FUNCTION "ROLL_PB25" : Void
{ S7_Optimized_Access := 'TRUE' }
VERSION : 0.1
VAR_TEMP
    r : Bool;
    a1 : Word;
    a2 : Word;
    activeDataBlock : Int;
    comparisonResults : Array[0..14] of Bool;
END_VAR
BEGIN
    #r := FALSE;
    #a1 := W#16#0000;
    #a2 := W#16#0000;
    #activeDataBlock := 0;
    // PB25, STEP 5 network 1
    #activeDataBlock := 15;
    // PB25, STEP 5 network 2
    #a2 := #a1;
    #a1 := "ROLL_GetM"(FirstByte := 5, Width := 8);
    #a2 := #a1;
    #a1 := W#16#0000;
    #comparisonResults[0] := (WORD_TO_INT(#a2) <> WORD_TO_INT(#a1));
    #r := #comparisonResults[0];
    "ROLL_State".M[87, 0] := #r;
    // PB25, STEP 5 network 3
    #a2 := #a1;
    #a1 := "ROLL_GetM"(FirstByte := 6, Width := 8);
    #a2 := #a1;
    #a1 := W#16#0000;
    #comparisonResults[1] := (WORD_TO_INT(#a2) <> WORD_TO_INT(#a1));
    #r := #comparisonResults[1];
    "ROLL_State".M[87, 1] := #r;
    // PB25, STEP 5 network 4
    #a2 := #a1;
    #a1 := "ROLL_GetM"(FirstByte := 7, Width := 8);
    #a2 := #a1;
    #a1 := W#16#0000;
    #comparisonResults[2] := (WORD_TO_INT(#a2) <> WORD_TO_INT(#a1));
    #r := #comparisonResults[2];
    "ROLL_State".M[87, 2] := #r;
    // PB25, STEP 5 network 5
    #a2 := #a1;
    #a1 := "ROLL_GetM"(FirstByte := 8, Width := 8);
    #a2 := #a1;
    #a1 := W#16#0000;
    #comparisonResults[3] := (WORD_TO_INT(#a2) <> WORD_TO_INT(#a1));
    #r := #comparisonResults[3];
    "ROLL_State".M[87, 3] := #r;
    // PB25, STEP 5 network 6
    #a2 := #a1;
    #a1 := "ROLL_GetM"(FirstByte := 9, Width := 8);
    #a2 := #a1;
    #a1 := W#16#0000;
    #comparisonResults[4] := (WORD_TO_INT(#a2) <> WORD_TO_INT(#a1));
    #r := #comparisonResults[4];
    "ROLL_State".M[87, 4] := #r;
    // PB25, STEP 5 network 7
    #a2 := #a1;
    #a1 := "ROLL_GetM"(FirstByte := 10, Width := 8);
    #a2 := #a1;
    #a1 := W#16#0000;
    #comparisonResults[5] := (WORD_TO_INT(#a2) <> WORD_TO_INT(#a1));
    #r := #comparisonResults[5];
    "ROLL_State".M[87, 5] := #r;
    // PB25, STEP 5 network 8
    #a2 := #a1;
    #a1 := "ROLL_GetM"(FirstByte := 11, Width := 8);
    #a2 := #a1;
    #a1 := W#16#0000;
    #comparisonResults[6] := (WORD_TO_INT(#a2) <> WORD_TO_INT(#a1));
    #r := #comparisonResults[6];
    "ROLL_State".M[87, 6] := #r;
    // PB25, STEP 5 network 9
    #a2 := #a1;
    #a1 := "ROLL_GetM"(FirstByte := 12, Width := 8);
    #a2 := #a1;
    #a1 := W#16#0000;
    #comparisonResults[7] := (WORD_TO_INT(#a2) <> WORD_TO_INT(#a1));
    #r := #comparisonResults[7];
    "ROLL_State".M[87, 7] := #r;
    // PB25, STEP 5 network 10
    #a2 := #a1;
    #a1 := "ROLL_GetM"(FirstByte := 13, Width := 8);
    #a2 := #a1;
    #a1 := W#16#0000;
    #comparisonResults[8] := (WORD_TO_INT(#a2) <> WORD_TO_INT(#a1));
    #r := #comparisonResults[8];
    "ROLL_State".M[88, 0] := #r;
    // PB25, STEP 5 network 11
    #a2 := #a1;
    #a1 := "ROLL_GetM"(FirstByte := 14, Width := 8);
    #a2 := #a1;
    #a1 := W#16#0000;
    #comparisonResults[9] := (WORD_TO_INT(#a2) <> WORD_TO_INT(#a1));
    #r := #comparisonResults[9];
    "ROLL_State".M[88, 1] := #r;
    // PB25, STEP 5 network 12
    #a2 := #a1;
    #a1 := "ROLL_GetM"(FirstByte := 15, Width := 8);
    #a2 := #a1;
    #a1 := W#16#0000;
    #comparisonResults[10] := (WORD_TO_INT(#a2) <> WORD_TO_INT(#a1));
    #r := #comparisonResults[10];
    "ROLL_State".M[88, 2] := #r;
    // PB25, STEP 5 network 13
    #a2 := #a1;
    #a1 := "ROLL_GetM"(FirstByte := 16, Width := 8);
    #a2 := #a1;
    #a1 := W#16#0000;
    #comparisonResults[11] := (WORD_TO_INT(#a2) <> WORD_TO_INT(#a1));
    #r := #comparisonResults[11];
    "ROLL_State".M[88, 3] := #r;
    // PB25, STEP 5 network 14
    #a2 := #a1;
    #a1 := "ROLL_GetM"(FirstByte := 17, Width := 8);
    #a2 := #a1;
    #a1 := W#16#0000;
    #comparisonResults[12] := (WORD_TO_INT(#a2) <> WORD_TO_INT(#a1));
    #r := #comparisonResults[12];
    "ROLL_State".M[88, 4] := #r;
    // PB25, STEP 5 network 15
    #a2 := #a1;
    #a1 := "ROLL_GetM"(FirstByte := 18, Width := 8);
    #a2 := #a1;
    #a1 := W#16#0000;
    #comparisonResults[13] := (WORD_TO_INT(#a2) <> WORD_TO_INT(#a1));
    #r := #comparisonResults[13];
    "ROLL_State".M[88, 5] := #r;
    // PB25, STEP 5 network 16
    #a2 := #a1;
    #a1 := "ROLL_GetM"(FirstByte := 19, Width := 8);
    #a2 := #a1;
    #a1 := W#16#0000;
    #comparisonResults[14] := (WORD_TO_INT(#a2) <> WORD_TO_INT(#a1));
    #r := #comparisonResults[14];
    "ROLL_State".M[88, 6] := #r;
    // PB25, STEP 5 network 17
    #r := ("ROLL_State".M[87, 0] OR "ROLL_State".M[87, 1] OR "ROLL_State".M[87, 2] OR "ROLL_State".M[87, 3] OR "ROLL_State".M[87, 4] OR "ROLL_State".M[87, 5] OR "ROLL_State".M[87, 6] OR "ROLL_State".M[87, 7] OR "ROLL_State".M[88, 0] OR "ROLL_State".M[88, 1] OR "ROLL_State".M[88, 2] OR "ROLL_State".M[88, 3] OR "ROLL_State".M[88, 4] OR "ROLL_State".M[88, 5] OR "ROLL_State".M[88, 6]);
    "ROLL_State".M[88, 7] := #r;
    // PB25, STEP 5 network 18
    #r := ("ROLL_IO".Input[1, 2] OR "ROLL_State".M[88, 7]);
    "ROLL_IO".Output[16, 4] := #r;
    // PB25, STEP 5 network 19
    #r := (("ROLL_State".M[3, 6] AND "ROLL_State".M[31, 6]) OR "ROLL_IO".Input[1, 2]);
    "ROLL_IO".Output[16, 5] := #r;
    // PB25, STEP 5 network 20
    #r := ("ROLL_IO".Input[1, 2] OR "ROLL_IO".Input[3, 4]);
    "ROLL_IO".Output[16, 0] := #r;
    // PB25, STEP 5 network 21
    #r := (((NOT "ROLL_State".M[31, 5]) AND "ROLL_State".M[28, 4]) OR ("ROLL_State".M[3, 6] AND "ROLL_State".M[74, 0]) OR "ROLL_IO".Input[1, 2]);
    "ROLL_IO".Output[16, 2] := #r;
    // PB25, STEP 5 network 22
    #r := (("ROLL_State".M[3, 6] AND "ROLL_State".M[31, 5]) OR "ROLL_IO".Input[1, 2] OR "ROLL_State".M[31, 4]);
    "ROLL_IO".Output[16, 3] := #r;
    // PB25, STEP 5 network 23
    #r := "ROLL_IO".Input[2, 0];
    "ROLL_IO".Output[19, 3] := #r;
    // PB25, STEP 5 network 24
    #r := (((("ROLL_IO".Input[14, 0] AND "ROLL_State".M[37, 1]) OR "ROLL_State".M[53, 6]) AND "ROLL_IO".Input[0, 2]) OR ("ROLL_IO".Input[0, 1] AND "ROLL_State".M[190, 6] AND "ROLL_State".M[20, 7]));
    IF #r THEN "ROLL_State".M[71, 5] := TRUE; END_IF;
    #r := (("ROLL_IO".Input[0, 1] AND "ROLL_State".M[190, 5] AND "ROLL_State".M[20, 7]) OR ("ROLL_IO".Input[0, 2] AND "ROLL_State".M[37, 2]));
    IF #r THEN "ROLL_State".M[71, 5] := FALSE; END_IF;
    #r := "ROLL_State".M[71, 5];
    "ROLL_IO".Output[17, 7] := #r;
    // PB25, STEP 5 network 25
    RETURN;
END_FUNCTION

FUNCTION "ROLL_PB50" : Void
{ S7_Optimized_Access := 'TRUE' }
VERSION : 0.1
VAR_TEMP
    r : Bool;
    a1 : Word;
    a2 : Word;
    activeDataBlock : Int;
    comparisonResults : Array[0..0] of Bool;
END_VAR
BEGIN
    #r := FALSE;
    #a1 := W#16#0000;
    #a2 := W#16#0000;
    #activeDataBlock := 0;
    // PB50, STEP 5 network 1
    #activeDataBlock := 15;
    // PB50, STEP 5 network 2
    #r := "ROLL_State".M[0, 1];
    IF #r THEN "ROLL_State".M[0, 2] := FALSE; END_IF;
    // PB50, STEP 5 network 3
    #a2 := #a1;
    #a1 := W#16#2008;
    #r := ((NOT "ROLL_State".M[0, 1]) AND "ROLL_IO".Input[3, 0]);
    "ROLL_TimerOp"(Number := 11, Operation := 0, Signal := #r, Preset := #a1);
    // PB50, STEP 5 network 4
    #a2 := #a1;
    #a1 := W#16#1020;
    #r := "ROLL_State".M[29, 0];
    "ROLL_TimerOp"(Number := 13, Operation := 0, Signal := #r, Preset := #a1);
    // PB50, STEP 5 network 5
    RETURN;
END_FUNCTION

FUNCTION "ROLL_PB51" : Void
{ S7_Optimized_Access := 'TRUE' }
VERSION : 0.1
VAR_TEMP
    r : Bool;
    a1 : Word;
    a2 : Word;
    activeDataBlock : Int;
    comparisonResults : Array[0..0] of Bool;
END_VAR
BEGIN
    #r := FALSE;
    #a1 := W#16#0000;
    #a2 := W#16#0000;
    #activeDataBlock := 0;
    // PB51, STEP 5 network 1
    #a2 := #a1;
    #a1 := W#16#2060;
    #r := "ROLL_IO".Output[24, 0];
    "ROLL_TimerOp"(Number := 15, Operation := 0, Signal := #r, Preset := #a1);
    // PB51, STEP 5 network 2
    #a2 := #a1;
    #a1 := W#16#3360;
    #r := ((NOT "ROLL_IO".Input[5, 6]) AND "ROLL_State".M[31, 5]);
    "ROLL_TimerOp"(Number := 16, Operation := 0, Signal := #r, Preset := #a1);
    // PB51, STEP 5 network 3
    #a2 := #a1;
    #a1 := W#16#1010;
    #r := "ROLL_State".M[37, 5];
    "ROLL_TimerOp"(Number := 18, Operation := 0, Signal := #r, Preset := #a1);
    // PB51, STEP 5 network 4
    #a2 := #a1;
    #a1 := W#16#2015;
    #r := (((NOT "ROLL_IO".Input[124, 1]) AND "ROLL_IO".Output[112, 1]) OR ((NOT "ROLL_IO".Input[124, 2]) AND "ROLL_IO".Output[112, 2]));
    "ROLL_TimerOp"(Number := 19, Operation := 0, Signal := #r, Preset := #a1);
    // PB51, STEP 5 network 5
    #a2 := #a1;
    #a1 := W#16#1010;
    #r := (("ROLL_IO".Input[123, 4] OR "ROLL_IO".Input[123, 5]) AND "ROLL_IO".Output[112, 0]);
    "ROLL_TimerOp"(Number := 20, Operation := 0, Signal := #r, Preset := #a1);
    // PB51, STEP 5 network 6
    #a2 := #a1;
    #a1 := W#16#1050;
    #r := "ROLL_IO".Input[123, 4];
    "ROLL_TimerOp"(Number := 21, Operation := 0, Signal := #r, Preset := #a1);
    // PB51, STEP 5 network 7
    #a2 := #a1;
    #a1 := W#16#2005;
    #r := ("ROLL_IO".Input[125, 0] AND "ROLL_IO".Input[125, 1]);
    "ROLL_TimerOp"(Number := 95, Operation := 0, Signal := #r, Preset := #a1);
    // PB51, STEP 5 network 8
    RETURN;
END_FUNCTION

FUNCTION "ROLL_PB52" : Void
{ S7_Optimized_Access := 'TRUE' }
VERSION : 0.1
VAR_TEMP
    r : Bool;
    a1 : Word;
    a2 : Word;
    activeDataBlock : Int;
    comparisonResults : Array[0..0] of Bool;
END_VAR
BEGIN
    #r := FALSE;
    #a1 := W#16#0000;
    #a2 := W#16#0000;
    #activeDataBlock := 0;
    // PB52, STEP 5 network 1
    #activeDataBlock := 15;
    // PB52, STEP 5 network 2
    #a2 := #a1;
    #a1 := "ROLL_GetDW"(DbNumber := #activeDataBlock, Index := 17);
    #r := ((NOT "ROLL_IO".Input[5, 5]) AND (NOT "ROLL_State".M[6, 3]) AND "ROLL_IO".Input[3, 1] AND "ROLL_State".M[4, 1] AND "ROLL_State".M[40, 5]);
    "ROLL_TimerOp"(Number := 17, Operation := 0, Signal := #r, Preset := #a1);
    // PB52, STEP 5 network 3
    #a2 := #a1;
    #a1 := "ROLL_GetDW"(DbNumber := #activeDataBlock, Index := 31);
    #r := ((NOT "ROLL_IO".Input[5, 3]) AND (NOT "ROLL_State".M[6, 1]) AND "ROLL_IO".Input[3, 1] AND "ROLL_State".M[4, 1]);
    "ROLL_TimerOp"(Number := 31, Operation := 0, Signal := #r, Preset := #a1);
    // PB52, STEP 5 network 4
    #a2 := #a1;
    #a1 := "ROLL_GetDW"(DbNumber := #activeDataBlock, Index := 32);
    #r := ((NOT "ROLL_IO".Input[6, 0]) AND (NOT "ROLL_State".M[6, 4]) AND "ROLL_IO".Input[3, 1] AND "ROLL_State".M[4, 1]);
    "ROLL_TimerOp"(Number := 32, Operation := 0, Signal := #r, Preset := #a1);
    // PB52, STEP 5 network 5
    #a2 := #a1;
    #a1 := "ROLL_GetDW"(DbNumber := #activeDataBlock, Index := 33);
    #r := ((NOT "ROLL_IO".Input[6, 2]) AND (NOT "ROLL_State".M[6, 5]) AND "ROLL_IO".Input[3, 1] AND "ROLL_State".M[4, 1]);
    "ROLL_TimerOp"(Number := 33, Operation := 0, Signal := #r, Preset := #a1);
    // PB52, STEP 5 network 6
    #a2 := #a1;
    #a1 := W#16#3030;
    #r := ((NOT "ROLL_State".M[0, 4]) AND (NOT "ROLL_State".M[6, 7]) AND "ROLL_IO".Input[3, 1] AND "ROLL_State".M[4, 1]);
    "ROLL_TimerOp"(Number := 35, Operation := 0, Signal := #r, Preset := #a1);
    // PB52, STEP 5 network 7
    #a2 := #a1;
    #a1 := W#16#3030;
    #r := ((NOT "ROLL_State".M[0, 4]) AND (NOT "ROLL_State".M[7, 0]) AND "ROLL_IO".Input[3, 1] AND "ROLL_State".M[4, 1]);
    "ROLL_TimerOp"(Number := 36, Operation := 0, Signal := #r, Preset := #a1);
    // PB52, STEP 5 network 8
    #a2 := #a1;
    #a1 := W#16#3030;
    #r := ((NOT "ROLL_State".M[0, 4]) AND (NOT "ROLL_State".M[7, 1]) AND "ROLL_IO".Input[3, 1] AND "ROLL_State".M[4, 1]);
    "ROLL_TimerOp"(Number := 37, Operation := 0, Signal := #r, Preset := #a1);
    // PB52, STEP 5 network 9
    #a2 := #a1;
    #a1 := W#16#3030;
    #r := ((NOT "ROLL_State".M[0, 4]) AND (NOT "ROLL_State".M[7, 2]) AND "ROLL_IO".Input[3, 1] AND "ROLL_State".M[4, 1]);
    "ROLL_TimerOp"(Number := 38, Operation := 0, Signal := #r, Preset := #a1);
    // PB52, STEP 5 network 10
    #a2 := #a1;
    #a1 := W#16#1005;
    #r := "ROLL_IO".Input[123, 1];
    "ROLL_TimerOp"(Number := 45, Operation := 0, Signal := #r, Preset := #a1);
    // PB52, STEP 5 network 11
    #a2 := #a1;
    #a1 := "ROLL_GetDW"(DbNumber := #activeDataBlock, Index := 58);
    #r := ("ROLL_IO".Input[3, 1] AND "ROLL_State".M[3, 6]);
    "ROLL_TimerOp"(Number := 58, Operation := 1, Signal := #r, Preset := #a1);
    #a2 := #a1;
    #a1 := "ROLL_GetDW"(DbNumber := #activeDataBlock, Index := 59);
    #r := ("ROLL_State".M[3, 6] AND "ROLL_State".S5Timers[58].Q);
    "ROLL_TimerOp"(Number := 59, Operation := 1, Signal := #r, Preset := #a1);
    // PB52, STEP 5 network 12
    #a2 := #a1;
    #a1 := "ROLL_GetDW"(DbNumber := #activeDataBlock, Index := 63);
    #r := (NOT "ROLL_State".S5Timers[62].Q);
    "ROLL_TimerOp"(Number := 63, Operation := 0, Signal := #r, Preset := #a1);
    #a2 := #a1;
    #a1 := "ROLL_GetDW"(DbNumber := #activeDataBlock, Index := 62);
    #r := "ROLL_State".S5Timers[63].Q;
    "ROLL_TimerOp"(Number := 62, Operation := 1, Signal := #r, Preset := #a1);
    #r := ((NOT "ROLL_State".M[103, 0]) AND (NOT "ROLL_State".M[103, 3]) AND (NOT "ROLL_State".M[103, 4]) AND (NOT "ROLL_State".S5Timers[119].Q));
    "ROLL_TimerOp"(Number := 62, Operation := 2, Signal := #r, Preset := #a1);
    // PB52, STEP 5 network 13
    #a2 := #a1;
    #a1 := W#16#2010;
    #r := "ROLL_IO".Input[5, 3];
    "ROLL_TimerOp"(Number := 70, Operation := 1, Signal := #r, Preset := #a1);
    // PB52, STEP 5 network 14
    #a2 := #a1;
    #a1 := W#16#2010;
    #r := "ROLL_IO".Input[6, 2];
    "ROLL_TimerOp"(Number := 72, Operation := 1, Signal := #r, Preset := #a1);
    // PB52, STEP 5 network 15
    #a2 := #a1;
    #a1 := "ROLL_GetDW"(DbNumber := #activeDataBlock, Index := 85);
    #r := "ROLL_State".M[41, 0];
    "ROLL_TimerOp"(Number := 85, Operation := 1, Signal := #r, Preset := #a1);
    // PB52, STEP 5 network 16
    RETURN;
END_FUNCTION
